ABB RobotStudio station: Práctica4_inicio.rspag

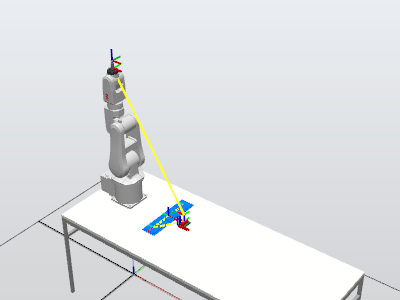
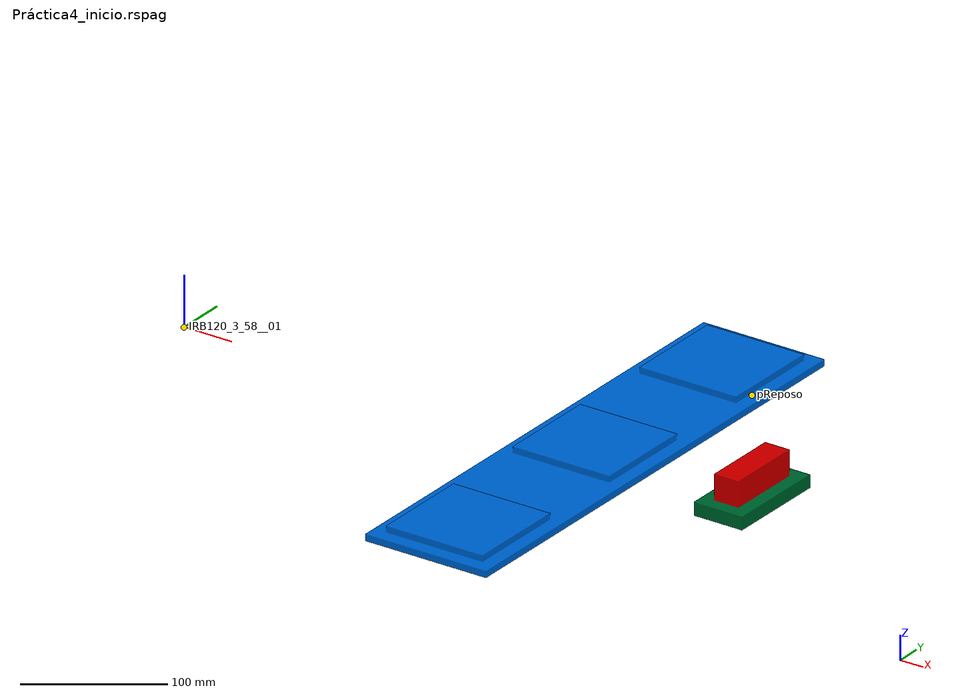
[picture v1: parts stored in the station drawn from their meshes, with robot base, taught points and paths (robot models come from the ABB library and are not in the file)]
--- station ---
Station Práctica3_inicio (saved by RobotStudio 25.2.11220.0)
Controller Controlador2, task T_ROB1: task frame (RAPID world) sits at (0, 0, 670) mm in the station
Controller Controlador2
  mechanical unit ROB_1: IRB120_3_58__01, 6 joints, base frame (0, 0, 0) mm
Layout (positions relative to the parent item):
  - TVentosa [mechanism] at (-70, 0, 1604) mm
      TCP TVentosa at (0, 0, 51.19) mm
      links: Mi_herramienta
  - LogicGate [smart component, from Components\LogicGate.rslib]
      properties: Operator=NOT; Delay=0
  - LogicGate_2 [smart component, from Components\LogicGate.rslib]
      properties: Operator=AND; Delay=0
  - IRB120_3_58__01 [mechanism, from %ABB.RobotStudio.Models.IRB120%\IRB120_3_58_G_01.rslib] at (0, 0, 670) mm; joint values [0, 0, -1.5708, 0, 0, 0] (rad or m)
  - table [part, from Libraries\e293a11e-ed86-4237-866f-a9bf8f4bd145table.rslib] at (-225, 300, 670) mm, rotated rx 0 ry 0 rz -90 deg
  - SimulationEvents [smart component, from Components\SimulationEvents.rslib]
  - Base0 [part], size 40 x 80 x 10 mm
  - Base [part], size 100 x 400 x 5 mm
  - Base1 [part], size 80 x 80 x 5 mm
  - Base2 [part], size 80 x 80 x 5 mm
  - Base3 [part], size 80 x 80 x 5 mm
  - Pieza [part] at (470, 0, 700) mm, rotated rx 180 ry 0 rz -90 deg, size 60 x 20 x 20 mm
  - CollisionSensor [smart component, from Components\CollisionSensor.rslib]
      properties: Object1=TVentosa; Object2=(none); NearMiss=0.001; Part1=(none); Part2=(none); CollisionType=0
  - Detacher [smart component, from Components\Detacher.rslib]
      properties: Child=(none); KeepPosition=true
  - Attacher [smart component, from Components\Attacher.rslib]
      properties: Parent=TVentosa; Flange=0; Child=(none); Mount=false; Offset=[0 0 0]; Orientation=[0 0 0]
  - Source [smart component, from Components\Source.rslib]
      properties: Source=Pieza; Copy=(none); Parent=(none); Position=[0.47 0 0.7]; Orientation=[3.14159265358979 0 -1.5707963267949]; Transient=true; PhysicsBehavior=0
Attachment: TVentosa is attached to IRB120_3_58__01 / Link6
Attachment: Base1 is attached to Base
Attachment: Base2 is attached to Base
Attachment: Base3 is attached to Base
Attachment: Pieza is attached to Base0
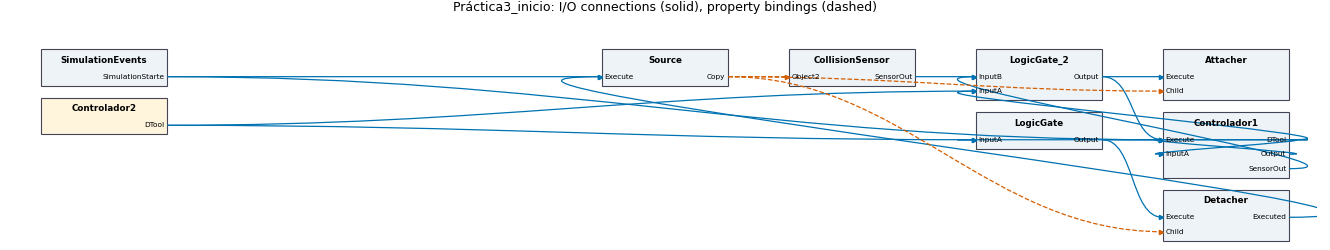
Station logic (signal -> signal, property => property):
  Controlador1.DTool -> Attacher.Execute
  Controlador1.DTool -> LogicGate_2.InputA
  LogicGate_2.Output -> Detacher.Execute
  Controlador1.DTool -> LogicGate.InputA
  LogicGate.Output -> Detacher.Execute
  CollisionSensor.SensorOut -> LogicGate_2.InputB
  Controlador1.DTool -> LogicGate_2.InputA
  LogicGate_2.Output -> Attacher.Execute
  SimulationEvents.SimulationStarted -> Source.Execute
  Controlador2.DTool -> LogicGate_2.InputA
  CollisionSensor.SensorOut -> LogicGate_2.InputB
  LogicGate_2.Output -> Attacher.Execute
  Controlador2.DTool -> LogicGate.InputA
  LogicGate.Output -> Detacher.Execute
  SimulationEvents.SimulationStarted -> Source.Execute
  Detacher.Executed -> Source.Execute
  Source.Copy => Attacher.Child
  Source.Copy => CollisionSensor.Object2
  Source.Copy => Detacher.Child
Targets, tools, work objects and paths stored in the station and not in the controller backup, written as RAPID:
! task T_ROB1
MODULE Module1
  PROC Path_10()
    MoveAbsJ Jhome,v1000,z100,TVentosa\WObj:=WO_Base;
    MoveJ pReposo,v1000,z100,TVentosa\WObj:=WO_Pieza;
    MoveJ pRecoger,v1000,z100,TVentosa\WObj:=WO_Pieza;
    MoveJ pBase1,v1000,z100,TVentosa\WObj:=WO_Base;
    MoveJ pBase2,v1000,z100,TVentosa\WObj:=WO_Base;
    MoveJ pBase3,v1000,z100,TVentosa\WObj:=WO_Base;
  ENDPROC
ENDMODULE


--- Backups/Controlador2/RAPID/TASK1/PROGMOD/CalibData.mod ---
MODULE CalibData
    PERS tooldata TVentosa:=[TRUE,[[0,0,51.19],[1,0,0,0]],[0.1,[0,0,1],[1,0,0,0],0,0,0]];
    TASK PERS wobjdata WO_Base:=[FALSE,TRUE,"",[[450,-40,10],[1,0,0,0]],[[-110,40,0],[1,0,0,0]]];
    TASK PERS wobjdata WO_Pieza:=[FALSE,TRUE,"",[[450,-40,10],[1,0,0,0]],[[10,10,0],[1,0,0,0]]];
ENDMODULE

--- Backups/Controlador2/RAPID/TASK1/PROGMOD/Module1.mod ---
MODULE Module1
    CONST jointtarget Jhome:=[[0,0,-90,0,0,0],[9E9,9E9,9E9,9E9,9E9,9E9]];
    CONST robtarget pReposo:=[[10,30,70],[0,0,1,0],[0,0,0,0],[9E9,9E9,9E9,9E9,9E9,9E9]];
    CONST robtarget pRecoger:=[[10,30,20],[0,0,1,0],[0,0,0,0],[9E9,9E9,9E9,9E9,9E9,9E9]];
    CONST robtarget pBase1:=[[0,-150,0],[0,-0.707106781,0.707106781,0],[0,0,-1,0],[9E9,9E9,9E9,9E9,9E9,9E9]];
    CONST robtarget pBase2:=[[0,0,0],[0,-0.707106781,0.707106781,0],[0,0,-1,0],[9E9,9E9,9E9,9E9,9E9,9E9]];
    CONST robtarget pBase3:=[[0,150,0],[0,-0.707106781,0.707106781,0],[0,0,-1,0],[9E9,9E9,9E9,9E9,9E9,9E9]];
    CONST num hPieza:=20;
    VAR num altura1;
    VAR num altura2;
    VAR num altura3;
    VAR num torre;

    PROC Initialize()
        altura1:=hPieza;
        altura2:=hPieza;
        altura3:=hPieza;
    ENDPROC

    PROC Pick(robtarget punto)
        MoveJ Offs(punto,0,0,50),v100,z10,TVentosa\WObj:=WO_Pieza;
        MoveL punto,v50,fine,TVentosa\WObj:=WO_Pieza;
        SetDO DTool,1;
        MoveL Offs(punto,0,0,50),v100,z10,TVentosa\WObj:=WO_Pieza;
    ENDPROC

    PROC Place(robtarget punto, VAR num altura)
        MoveJ Offs(punto,0,0,50+altura),v100,z10,TVentosa\WObj:=WO_Base;
        MoveL Offs(punto,0,0,altura),v50,fine,TVentosa\WObj:=WO_Base;
        SetDO DTool,0;
        MoveL Offs(punto,0,0,50+altura),v100,z10,TVentosa\WObj:=WO_Base;
        altura:=altura+hPieza;
    ENDPROC

    PROC main()
        Initialize;
        MoveAbsJ Jhome,v1000,fine,TVentosa;
        MoveJ pReposo,v1000,z100,TVentosa\WObj:=WO_Pieza;
        FOR i FROM 1 TO 10 DO
            TPReadNum torre,"Elige torre (1-3):";
            Pick pRecoger;
            IF torre=1 THEN
                Place pBase1,altura1;
            ELSEIF torre=2 THEN
                Place pBase2,altura2;
            ELSEIF torre=3 THEN
                Place pBase3,altura3;
            ENDIF
        ENDFOR
        MoveAbsJ Jhome,v1000,fine,TVentosa;
    ENDPROC
ENDMODULE

--- Backups/Controlador2/SYSPAR/EIO.cfg ---
EIO:CFG_1.0:6:1::
#
EIO_SIGNAL:

      -Name "DTool" -SignalType "DO"
